(* IEC 61131-3 sources: kns-port-domestic/tools/port_metrics_tests/fixtures/adapted/src/POUs/FB_Base, 1 file *)

(* ---- FB_Base.decl.st ---- *)
// PORT: [oop] база больше не наследуется
FUNCTION_BLOCK FB_Base
VAR_OUTPUT
    xFault : BOOL;
END_VAR
